SUBAPPLICATION IN_UP (* Subapplication Type *)
  (* Standard: 61499-2 *)
  (* Version 1.0, 2023-02-06, franz *)
  IMPORT BlinkMarine::io::DI::PKP_2200_LI_DI::Invalid;
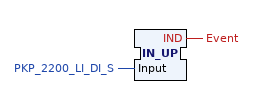
  EVENT_OUTPUT
    IND;
  END_EVENT
  VAR_INPUT
    Input : BlinkMarine::io::DI::PKP_2200_LI_DI_S := Invalid;
  END_VAR
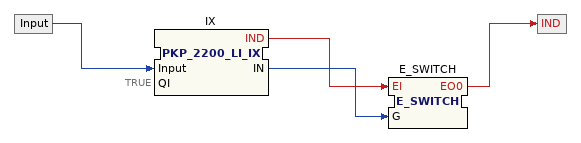
  FBS
    E_SWITCH : E_SWITCH;
    IX : BlinkMarine::io::DI::PKP_2200_LI_IX(QI := TRUE);
  END_FBS
  EVENT_CONNECTIONS
    IX.IND TO E_SWITCH.EI;
    E_SWITCH.EO0 TO IND;
  END_CONNECTIONS
  DATA_CONNECTIONS
    Input TO IX.Input;
    IX.IN TO E_SWITCH.G;
  END_CONNECTIONS
END_SUBAPPLICATION
